(* PLC project PumpStation, Demo Demo 1 *)
(* stored: creationDateTime 2026-01-01T00:00:00 *)

PROGRAM PumpControl
  VAR
    Pressure AT %IW0 : INT;
  END_VAR

IF Pressure > Setpoint THEN
    ReliefValve := TRUE;
ELSE
    ReliefValve := FALSE;
END_IF;
PumpRun := PumpSpeed > 0 AND PumpSpeed <= SpeedLimit;
Runtime := Runtime + 1;
IF Runtime > 4000000 THEN
    PumpRun := FALSE;
END_IF;
END_PROGRAM

PROGRAM Panel

(* LD diagram, written out as Structured Text *)
END_PROGRAM

CONFIGURATION Config
  RESOURCE Res ON PLC
    VAR_GLOBAL
      PumpSpeed AT %MW0 : INT;
      SpeedLimit AT %MW1 : INT := 1500;
      Setpoint AT %MW10 : INT;  (* pressure setpoint kPa *)
      ReliefValve AT %QX0.1 : BOOL;
      PumpRun AT %QX0.0 : BOOL;
      Runtime : DINT;
      Recipe AT %MW30 : ARRAY[0..3] OF REAL;
    END_VAR
  END_RESOURCE
END_CONFIGURATION
